Fanuc KAREL source: KT00068.KL

PROGRAM KT00068
%NOLOCKGROUP
VAR
  I1: INTEGER
  R2: REAL
  OUT: REAL
BEGIN
  I1 = 2
    R2 = 3.0
  OUT = I1 * R2
END KT00068
